RoboDK station: ROBODK_DOBOT.rdk

Station New Station (saved by RoboDK 6.0.1). Poses are relative to the parent item; angles as X-Y-Z fixed-axis rotations.
